(* IEC 61131-3 sources: Caravan/Archiv/12-04-19/Stations/MachineControl/MachineControl/Class/VaranManager (part 3) *)

#ifndef VARAN_TIME_MEASUREMENT_DEACTIVATE
        if pMultiVaran^.udVersion >= VM_MULTIVARAN_VERSION_FULL_PAYLOAD_AVAILABLE then
          //save max response time
          if ( p_node_info^^.uiResponseTimeMax > s_VaranTimes.ud_MaxResponseTime ) then

            s_VaranTimes.ud_MaxResponseTime := p_node_info^^.uiResponseTimeMax;

            //set T3 (no command executed before isochronous task)
            s_ManagerControlData.ud_MaxTimeCmdExecution := s_ManagerControlData.ud_IsoStartPoint -
                                  (2*( ( ( 276 * VM_TIMEOUT_ONE_BYTE )			//max 128 read/write befehl
                                    + s_VaranTimes.ud_MaxResponseTime       //The Manager need 2 Commands before he is free ( Prefetch + actual Command), reason for the whole term multiple 2
                                    )                                       //minimize the Jitter from the VARAN-BUS
                                    * ( VM_ALLOWED_RETRIES + 1 ))
                                  );

            //if time is neg set to 0
            if ( s_ManagerControlData.ud_MaxTimeCmdExecution$DINT < 0 ) then
              s_ManagerControlData.ud_MaxTimeCmdExecution := 0;
            end_if;

            // Write the data
            nodeProperty.udPropertyId    := VM_PROP_MAX_COMMAND_EXECUTION_TIME;
            nodeProperty.udPropertyValue := s_ManagerControlData.ud_MaxTimeCmdExecution;
            MULTI_VARAN_iSetNodeProperties( hNodeHandle           := vmNodeHandle
                                          , udPropertyCount       := 1
                                          , psPropertyValuePairs  := #nodeProperty
                                          );

          end_if;

        else
          //save max response time
          if ( p_node_info^^.uiResponseTimeMax > s_VaranTimes.ud_MaxResponseTime ) & p_ManagerStructure then

            s_VaranTimes.ud_MaxResponseTime := p_node_info^^.uiResponseTimeMax;

            //set T3 (no command executed before isochronous task)
            p_ManagerStructure^.uiMaxTimeCmdExecution := 	p_ManagerStructure^.uiIsoStartPoint -
                                  (2*( ( ( 276 * VM_TIMEOUT_ONE_BYTE )			//max 128 read/write befehl
                                    + s_VaranTimes.ud_MaxResponseTime       //The Manager need 2 Commands before he is free ( Prefetch + actual Command), reason for the whole term multiple 2
                                    )                                       //minimize the Jitter from the VARAN-BUS
                                    * ( VM_ALLOWED_RETRIES + 1 ))
                                  );

            //if time is neg set to 0
            if ( p_ManagerStructure^.uiMaxTimeCmdExecution$DINT < 0 ) then
              p_ManagerStructure^.uiMaxTimeCmdExecution := 0;
            end_if;
          end_if;
        end_if;
#endif

      else
        sd_retval := VM_CMD_ERROR_EMPTY_POINTER;
      end_if;

    elsif pVaran then  // if b_PayloadSupport then //----------------------------------------------------------------------------------------------------------

      //call OS - function to right device address
      sd_retval := VARAN_iGetNodeInfo	( uiManager	:= VaranManagerNr
                                      , pucNode	  := p_us_position_info
                                      , pNodeInfo	:= p_node_info
                                      );

      //look for an Error
      if ( sd_retval <> VARANMANAGER_OK ) then
        s_ErrorVaranManager.f_GetNodeInfo := SetVaranDOError( sd_Error 		  := sd_retval
                                                            , b_manager_off	:= FALSE
                                                            , b_log			    := FALSE
                                                            );
        return;
      end_if;

#ifndef VARAN_TIME_MEASUREMENT_DEACTIVATE
      //save max response time
      if ( p_node_info^^.uiResponseTimeMax > s_VaranTimes.ud_MaxResponseTime ) & p_ManagerStructure then

        s_VaranTimes.ud_MaxResponseTime := p_node_info^^.uiResponseTimeMax;

        //set T3 (no command executed before isochronous task)
        p_ManagerStructure^.uiMaxTimeCmdExecution := 	p_ManagerStructure^.uiIsoStartPoint -
                              (2*( ( ( 276 * VM_TIMEOUT_ONE_BYTE )			//max 128 read/write befehl
                                + s_VaranTimes.ud_MaxResponseTime       //The Manager need 2 Commands before he is free ( Prefetch + actual Command), reason for the whole term multiple 2
                                )                                       //minimize the Jitter from the VARAN-BUS
                                * ( VM_ALLOWED_RETRIES + 1 ))
                              );

        //if time is neg set to 0
        if ( p_ManagerStructure^.uiMaxTimeCmdExecution$DINT < 0 ) then
          p_ManagerStructure^.uiMaxTimeCmdExecution := 0;
        end_if;
      end_if;
#endif
    end_if;	  // if b_PayloadSupport then //----------------------------------------------------------------------------------------------------------

  else
    sd_retval := -101;
  end_if;

END_FUNCTION //VIRTUAL GLOBAL VaranManager::GetNodeInfo

//[#ENGLISH]
//=================================================================================================
//Function to get Varan Manager number
//=================================================================================================
//[clients]	VaranManagerNr		:R		:number of varan manager
//[members]	pVaran					:R		:pointer to varan os functions
//			s_VaranManagerSettings	:R		:structure for different varan settings
//[<sd_Manager_number]number of varan Manager
//[>p_varan]address of pointer to varan
FUNCTION VIRTUAL GLOBAL VaranManager::GetManagerNumber
  VAR_INPUT
    p_varan				    : ^pVoid;
  END_VAR
  VAR_OUTPUT
    ud_manager_number	:  UDINT;
  END_VAR

  //look if init was executed
  if ( s_VaranManagerSettings.us_InitCounter = 0 ) then
    bExternalInit := true;
    Init();
  end_if;

  //set pointer to varan functions
  p_varan^:= pVaran;

  //give back varan manager number
  ud_manager_number := VaranManagerNr.read();

END_FUNCTION //VIRTUAL GLOBAL VaranManager::GetManagerNumber

//[#ENGLISH]
//=================================================================================================
//Function to log faults in cyclic (to prevent an error 67)
//=================================================================================================
//[server]	State					:W		:State of class
//[members]	s_VaranManagerSettings	:W		:structure for different varan settings
FUNCTION  VaranManager::LogError
  VAR
    ud_reason	      : UDINT;
    b_SetError    	: BOOL;
  END_VAR

  ud_reason := 0;

  b_SetError := FALSE;

  //look which entry
  case ( State ) of
//**********************************************************************************************************************************************************
    _TimeSliceError:	//Log entry
#ifdef HWC_LogError
      HWC_LogError(this, "@06B8 (VaranManager::LogError) Timeslice Error! Manager is set off!");
#endif
      ud_reason := VM_ERROR_TIMESLICE;
      b_SetError := TRUE;

//**********************************************************************************************************************************************************
    _TimesliceErrorIRQ:	//Log entry
#ifdef HWC_LogError
      HWC_LogError(this, "@06C2 (VaranManager::LogError) Timeslice Error Interrupt, Manager is set off!");
#endif
      ud_reason := VM_ERROR_TIMESLICE_IRQ;
      b_SetError := TRUE;

//**********************************************************************************************************************************************************
    _WatchdogError:		//Log entry
#ifdef HWC_LogError
      HWC_LogError(this, "@06CC (VaranManager::LogError) Watchdog Error Interrupt, Manager is set off!");
#endif
      ud_reason := VM_ERROR_WATCHDOG;
      b_SetError := TRUE;

//**********************************************************************************************************************************************************
    _RequiredError:		//Log entry
#ifdef HWC_LogError
      HWC_LogError(this, "@06D6 (VaranManager::LogError) Required Module not ready, Manager is set off!");
#endif
      //b_SetError := FALSE;

//**********************************************************************************************************************************************************
    _DeviceError:		//Log entry
#ifdef HWC_LogError
      HWC_LogError(this, "@06E0 (VaranManager::LogError) Error on Device, Manager is set off!");
#endif
      ud_reason := VM_ERROR_DEVICE;
      b_SetError := TRUE;

//**********************************************************************************************************************************************************
    _CDIASRequiredError, _DIASRequiredError, _DiasError: //Log Entry
#ifdef HWC_LogError
      HWC_LogError(this, "@0024 (VaranManager::LogError) Required DIAS/CDIAS Module not ready, Manager is set off!");
#endif
      ud_reason   := VM_ERROR_DEVICE;
      b_SetError  := TRUE;
      State       := _RequiredError;

//**********************************************************************************************************************************************************
  else     //Unknown fault, log that an error occured
#ifdef HWC_LogValue1
    HWC_LogValue1(this, "@0025 (VaranManager::LogError) Unknown Fault (State = {0}), Manager is set off!", State);
#endif
  end_case;

  //reset log flag
  s_VaranManagerSettings.b_LogError := FALSE;

  //set Hw off
  To_HwControl.SetHardwareOff( e_error := State );

  //produce Varan Manager Error
  if ( b_SetError & PreventManagerError = 0) then

    if b_PayloadSupport & pMultiVaran^.udVersion >= VM_MULTIVARAN_VERSION_FULL_PAYLOAD_AVAILABLE  then
      MULTI_VARAN_iReportVaranError(diErrorNumber := ud_reason$DINT
                                  , hErrorNode    := vmNodeHandle);

    elsif pVaran & (pVaran^.udVersion >= 16#00001104 ) then
      VARAN_iSetManagerError( VaranManagerNr, ud_reason );
    end_if;
  end_if;

END_FUNCTION // VaranManager::LogError

//[#ENGLISH]
//=================================================================================================
//Function returns state of Varan manger class
//=================================================================================================
//[<e_state]error of varan manager
FUNCTION VIRTUAL GLOBAL VaranManager::GetManagerState
  VAR_OUTPUT
    e_state		  : t_e_VaranErrors;
  END_VAR

  e_state := State;

END_FUNCTION //VIRTUAL GLOBAL VaranManager::GetManagerState

//[#ENGLISH]
//=================================================================================================
//Function to add a multiple read/write register
//=================================================================================================
//[>p_us_position_info]pointer to position info( first byte is length)
//[>ud_dol_type] type of DOL list( 1=direct access, 2=IRQ, 3=realtime, 4=cyclic )
//[>p_ud_handle] pointer to variable to set right handle
//[>ud_address_read] Address of read data object
//[>ud_length_read] Length of read data object
//[>p_ud_data_read] pointer to variable to get pointer to data
//[>ud_address_write] Address of write data object
//[>ud_length_write] Length of write data object
//[>p_ud_data_write] pointer to variable to get pointer to data
//[>us_filter]filter number
//[>ui_number_of_slices]maximal number of slices
//[<sd_retval] 0=OK, negative=error (look lsl_st_varan.h)
FUNCTION GLOBAL VaranManager::AddMultipleRdWr
  VAR_INPUT
    p_us_position_info		: ^USINT;
    ud_dol_type				    :  UDINT;
    p_ud_handle				    : ^UDINT;
    ud_address_read			  :  UDINT;
    ud_length_read			  :  UDINT;
    p_ud_data_read			  : ^UDINT;
    ud_address_write		  :  UDINT;
    ud_length_write			  :  UDINT;
    p_ud_data_write			  : ^UDINT;
    us_filter				      :  USINT;
    ui_number_of_slices		:  UINT;
  END_VAR
  VAR_OUTPUT
    sd_retval				      :  DINT;
  END_VAR
  VAR
    ud_command			      :  UDINT;
    TempMem               :  UDINT;
  END_VAR

  //look if right OS - Version
  if ( _RTOSVersion >= 16#1194 ) & pVaran then

    //set command
    ud_command := VARAN_CMD_MULTIPLE_MEMORY_RW or ( us_filter shl 8 ) or ( ui_number_of_slices shl 16 );

    //look if we must execute Cyclic DOL list
    if ( ud_dol_type = VARAN_DOL_ASY ) then
      s_CyHandles.b_ExecuteDOL := TRUE;			//set flag to execut Dol list
    end_if;

    //Install Varan data object
    sd_retval := VARAN_iAddDOToDOL( uiManager     := VaranManagerNr
                                  , pucNode       := p_us_position_info
                                  , uiDOLType     := ud_dol_type
                                  , puiDOHandle   := p_ud_handle
                                  , uiCmd				  := ud_command
                                  , uiAddressRead := ud_address_read
                                  , uiLengthRead  := ud_length_read
                                  , pucRead       := p_ud_data_read
                                  , uiAddressWrite:= ud_address_write
                                  , uiLengthWrite := ud_length_write
                                  , pucWrite      := p_ud_data_write
                                  );

    //look if an error occured
    if ( sd_retval <> VARANMANAGER_OK ) then
      s_ErrorVaranManager.f_AddRdWrDO := SetVaranDOError( sd_Error      := sd_retval
                                                        , b_manager_off := TRUE
                                                        , b_log         := TRUE
                                                        );
    else
    //   32Byte (Header) +
    // + 13 Byte (Addr + Len +... --> See design spec appendix) +
    // + (1 Byte (Response) + n Byte) * slices (load data read) +
    // + n * slices Byte (load data write) +
    // + 0 to 3 Byte (compensate missalignment)
      TempMem := 32 + 13 + (1 + ud_length_read) * ui_number_of_slices + ud_length_write * ui_number_of_slices;
      if (TempMem MOD 4) then
        TempMem := TempMem + (4 - (TempMem MOD 4)); //increase memory, up to a value, which could be divided by 4
      end_if;

      if ud_dol_type = VARAN_DOL_ISO then
        DPRAM_Used.ISO_RdWr += TempMem;
        DOCounter.ISO_RdWr  += 1;
      else
        DPRAM_Used.ASY_RdWr += TempMem;
        DOCounter.ASY_RdWr  += 1;
      end_if;

      DPRAM_Used.Total      += TempMem;
      DOCounter.Total       += 1;
    end_if;
  else
    sd_retval := -100;	//Manager is off
  end_if;

END_FUNCTION //VIRTUAL GLOBAL VaranManager::AddMultipleRdWr

//[#ENGLISH]
//=================================================================================================
//Function to get an actual filter number
//=================================================================================================
//[<us_filter]number of filter
FUNCTION GLOBAL VaranManager::GetFilterNumber
  VAR_OUTPUT
    us_filter : USINT;
  END_VAR

  if ( s_VaranManagerSettings.us_FilterNumber <> 255 ) then
    //increment filter number
    s_VaranManagerSettings.us_FilterNumber += 1;
    us_filter := s_VaranManagerSettings.us_FilterNumber;
  else
    us_filter := 0;
  end_if;

END_FUNCTION //VIRTUAL GLOBAL VaranManager::GetFilterNumber

//[#ENGLISH]
//=================================================================================================
//Function to write a direct access data object
//=================================================================================================
//[members]	s_DirectAccessDO	:W/R	:structure for direct access
//[>p_us_position_info]pointer to position info( first byte is length)
//[>ud_address_read] Address of read data object
//[>ud_length_read] Length of read data object
//[>p_ud_data_read] pointer to variable to get pointer to data
//[>ud_address_write] Address of write data object
//[>ud_length_write] Length of write data object
//[>p_ud_data_write] pointer to variable to get pointer to data
//[>us_filter] number of filter
//[>us_slices] max number of slices
//[>p_handle]pointer to varan header
//[<sd_retval] 0=OK, negative=error (look lsl_st_varan.h)
FUNCTION GLOBAL VaranManager::MultipleRdWrDO
  VAR_INPUT
    p_us_position_info	: ^USINT;
    ud_address_read		  :  UDINT;
    ud_length_read		  :  UDINT;
    p_ud_data_read		  : ^UDINT;
    ud_address_write  	:  UDINT;
    ud_length_write		  :  UDINT;
    p_ud_data_write	  	: ^UDINT;
    us_filter			      :  USINT;
    us_slices			      :  USINT;
    p_handle			      : ^PLSL_VARANFRAME;
  END_VAR
  VAR_OUTPUT
    sd_retval		      	:  DINT;
  END_VAR

  //look if right OS - Version
  if ( _RTOSVersion >= 16#1194 ) then

    //clear direct access dol list
    sd_retval := ClearDOL( ud_dol_type := VARAN_DOL_DA );

    //look if an error occurs
    if ( sd_retval <> VARANMANAGER_OK ) then
      s_ErrorVaranManager.f_WrDO := SetVaranDOError	( sd_Error 	    := sd_retval
                                                    , b_manager_off	:= TRUE
                                                    , b_log			    := FALSE
                                                    );
      return;
    end_if;

    //add data object
    sd_retval := AddMultipleRdWr( p_us_position_info	:= p_us_position_info
                                , ud_dol_type			    := VARAN_DOL_DA
                                , p_ud_handle			    := p_handle$^UDINT
                                , ud_address_read		  := ud_address_read
                                , ud_length_read		  := ud_length_read
                                , p_ud_data_read		  := ( #p_ud_data_read )$^UDINT
                                , ud_address_write		:= ud_address_write
                                , ud_length_write		  := ud_length_write
                                , p_ud_data_write		  := ( #p_ud_data_write )$^UDINT
                                , us_filter				    := us_filter
                                , ui_number_of_slices	:= us_slices
                                );

    //look if an error occurs
    if ( sd_retval <> VARANMANAGER_OK ) then
      s_ErrorVaranManager.f_WrDO := SetVaranDOError	( sd_Error 		  := sd_retval
                                                    , b_manager_off	:= TRUE
                                                    , b_log			    := FALSE
                                                    );
      return;
    end_if;

    //set run status of data object on
    p_handle^^.ucCtrlStat 	        := VARAN_DO_SINGLE_RUN;

    //set number of allowed retries
    p_handle^^.ucRetrys	          	:= VM_ALLOWED_RETRIES;

    //set time for retry timeout
    p_handle^^.uiRetryTimeout       := VM_MAX_RETRY_TIMEOUT_MULTIPLE;

    //Execute dol
    sd_retval := ExecuteDOL( ud_dol_type := VARAN_DOL_DA );//or VARAN_DOL_EXECUTE_WAIT );

    //look if an error occurs
    if ( sd_retval <> VARANMANAGER_OK ) then
      s_ErrorVaranManager.f_WrDO := SetVaranDOError	( sd_Error 		  := sd_retval
                                                    , b_manager_off	:= TRUE
                                                    , b_log			    := FALSE
                                                    );
      return;
    end_if;

  else
    sd_retval := -100;	//Manager is off
  end_if;

END_FUNCTION //VIRTUAL GLOBAL VaranManager::MultipleRdWrDO

//[#ENGLISH]
//=================================================================================================
//Function to read SPI data
//=================================================================================================
//[>p_us_position_info]pointer to position info( first byte is length)
//[>ud_offset]offset in SPI flash
//[>ud_length]length of data (max. 128Byte)
//[>p_data]pointer to allocated memory for read data
//[<sd_retval] 0=OK, negative=error (look lsl_st_varan.h)
FUNCTION VIRTUAL GLOBAL VaranManager::ReadSPIData
  VAR_INPUT
    p_us_position_info	  : ^USINT;
    ud_offset		        	:  UDINT;
    ud_length		        	:  UDINT;
    p_data			        	: ^USINT;
  END_VAR
  VAR_OUTPUT
    sd_retval		          :  DINT;
  END_VAR
  VAR
    ud_sent_page	        :  UDINT;
    ud_NodeHandle         : UDINT;
    sPropertyValuePair    : LSL_PROPERTY_VALUE_PAIR;
  END_VAR

  //look if right OS - Version
  if ( _RTOSVersion >= 16#119F ) then

    if ( ud_length and VM_SPI_IDENT_LIST ) then
      ud_length     := ud_length and 16#7FFF_FFFF;
      ud_sent_page  := 16#FFFF_FFFF;   // = Read from the last page
    else
      ud_sent_page  := ud_offset / VM_SPI_PAGE_SIZE;
    end_if;

    //look for length
    if ( ud_length <= 0 | ud_length > 128 | p_data = NIL ) then
      sd_retval := -101;
      return;
    end_if;

    if b_PayloadSupport then
      // Get Node Handle
      sd_retval := MULTI_VARAN_iGetNodeHandle ( udManagerNumber := VaranManagerNr
                                              , pszHardwarePath := p_us_position_info
                                              , phNodeHandle    := #ud_NodeHandle
                                              );

      if sd_retval <> VARANMANAGER_OK then
        return;
      end_if;

      // set request
      sPropertyValuePair.udPropertyId     := ND_PROP_SPI_MASTER_REQUEST;
      sPropertyValuePair.udPropertyValue  := SPI_MASTER_REQ_SET;
      sd_retval := MULTI_VARAN_iSetNodeProperties ( hNodeHandle           := ud_NodeHandle
                                                  , udPropertyCount       := 1
                                                  , psPropertyValuePairs  := #sPropertyValuePair
                                                  );
      // look for an error
      if ( sd_retval <> VARANMANAGER_OK ) then
        return;
      end_if;

      // set right page
      sd_retval := MULTI_VARAN_iSpiMasterReadFlashPage( hNodeHandle           := ud_NodeHandle
                                                      , udPageNumber          := ud_sent_page
                                                      , udOffsetInPage        := ud_offset mod VM_SPI_PAGE_SIZE
                                                      , udReadLength          := ud_length
                                                      , bBlockUntilCompleted  := true
                                                      , pusData               := p_data
                                                      );
      //look for an error
      if ( sd_retval <> VARANMANAGER_OK ) then
        return;
      end_if;

      //clear request
      sPropertyValuePair.udPropertyId     := ND_PROP_SPI_MASTER_REQUEST;
      sPropertyValuePair.udPropertyValue  := SPI_MASTER_REQ_CLEARED;
      sd_retval := MULTI_VARAN_iSetNodeProperties ( hNodeHandle           := ud_NodeHandle
                                                  , udPropertyCount       := 1
                                                  , psPropertyValuePairs  := #sPropertyValuePair
                                                  );
    elsif pVaran then

      //set request
    sd_retval := VARAN_iSPIMasterSetRequest	( uiManager	:= VaranManagerNr
                                            , pucNode	  := p_us_position_info
                                            );

    //look for an error
    if ( sd_retval <> VARANMANAGER_OK ) then
      return;
    end_if;

    //set right page
    sd_retval := VARAN_iSPIMasterPageRead	( uiManager	:= VaranManagerNr
                                          , pucNode	  := p_us_position_info
                                          , uiPage	  := ud_sent_page
                                          );

    //look for an error
    if ( sd_retval <> VARANMANAGER_OK ) then
      return;
    end_if;

    ud_sent_page := ud_offset mod VM_SPI_PAGE_SIZE;

    //read data of page
    sd_retval := VARAN_iSPIMasterPageReadBuffer	( uiManager	:= VaranManagerNr
                                                , pucNode	  := p_us_position_info
                                                , uiOffset	:= ud_sent_page
                                                , uiLen		  := ud_length
                                                , puiPage	  := p_data
                                                );

    //look for an error
    if ( sd_retval <> VARANMANAGER_OK ) then
      return;
    end_if;

    //clear request
    sd_retval := VARAN_iSPIMasterClearRequest	( uiManager	:= VaranManagerNr
                                              , pucNode	  := p_us_position_info
                                              );
    end_if;

  else
    sd_retval := -100;
  end_if;

END_FUNCTION //VIRTUAL GLOBAL VaranManager::ReadSPIData

//[#ENGLISH]
//=================================================================================================
//Function add a foreign package request
//=================================================================================================
//[>p_us_position_info]pointer to position info( first byte is length)
//[>ud_dol_type] type of DOL list( 1=direct access, 2=IRQ, 3=realtime, 4=cyclic )
//[>p_ud_handle]pointer to variable to set right handle
//[>ud_address] Address of data object
//[<sd_retval] 0=OK, negative=error (look lsl_st_varan.h)
FUNCTION VIRTUAL GLOBAL VaranManager::AddForeignPackRequest
  VAR_INPUT
    p_us_position_info	: ^USINT;
    ud_dol_type		    	: UDINT;
    p_ud_handle			    : ^UDINT;
    ud_address			    : UDINT;
  END_VAR
  VAR_OUTPUT
    sd_retval		      	: DINT;
  END_VAR
  VAR
    ud_NodeHandle       : UDINT;
  END_VAR

  //look if we must execute Cyclic DOL list
  if ( ud_dol_type = VARAN_DOL_ASY ) then
    s_CyHandles.b_ExecuteDOL := TRUE;			//set flag to execut Dol list
  end_if;

  if b_PayloadSupport &
       pMultiVaran^.udVersion >= VM_MULTIVARAN_VERSION_FULL_PAYLOAD_AVAILABLE  then
    sd_retval := MULTI_VARAN_iGetNodeHandle ( udManagerNumber := VaranManagerNr
                                            , pszHardwarePath := p_DisablePath
                                            , phNodeHandle    := #ud_NodeHandle
                                            );

    // Return the ErrorCode
    if sd_retval then
      return;
    end_if;

    sd_retval := MULTI_VARAN_iAddDo(  phDoHandle                    := p_ud_handle
                                    , hNodeHandle                   := ud_NodeHandle
                                    , bDoRequired                   := 0
                                    , udDolType                     := ud_dol_type
                                    , udCommand                     := VARAN_CMD_FOREIGN_PACKET_REQ
                                    , udPriority                    := VM_PRIORITY_READ_DO
                                    , udPrescalerCounterThreshold   := 0
                                    , udPrescalerCounterStartValue  := 0
                                    , udReadOffset                  := VARAN_CLIENT_FP_SAFETY
                                    , udReadLength                  := VARAN_FPR_SAFETY_ID
                                    , udWriteOffset                 := 0
                                    , udWriteLength                 := 0
                                    , udFilter                      := 0
                                    , udSlices                      := 0
                                    , udWritePayloadType            := WR_PLD_TYPE_STANDARD
                                    );

  else
    // if there is no VARAN Interface available, we would crash at the call
    if pVaran = NIL then
      sd_retval := VARANMANAGER_DRIVER_NOT_EXISTS;
      return;
    end_if;

    //Install Varan data object
    sd_retval := VARAN_iAddDOToDOL	( uiManager			  := VaranManagerNr
                                    , pucNode			    := p_us_position_info
                                    , uiDOLType 		  := ud_dol_type + ( VARAN_DO_EXECUTE_FIFO_EMPTY shl 24 ) // in the highest byte we have the init value for the uc_CtrlStat Register
                                    , puiDOHandle		  := p_ud_handle
                                    , uiCmd				    := VARAN_CMD_FOREIGN_PACKET_REQ
                                    , uiAddressRead		:= ud_address + VARAN_CLIENT_FP_SAFETY
                                    , uiLengthRead		:= VARAN_FPR_SAFETY_ID
                                    , pucRead			    := NIL
                                    , uiAddressWrite	:= 0
                                    , uiLengthWrite		:= 0
                                    , pucWrite			  := NIL
                                    );
  end_if;

  //look if an error occured
  if ( sd_retval <> VARANMANAGER_OK ) then
    s_ErrorVaranManager.f_AddFoPaReq := SetVaranDOError ( sd_Error 		  := sd_retval
                                                        , b_manager_off	:= TRUE
                                                        , b_log			    := TRUE
                                                        );
  end_if;

  //look if an error occured
  if ( sd_retval <> VARANMANAGER_OK ) then
    s_ErrorVaranManager.f_AddFoPaReq := SetVaranDOError ( sd_Error 		  := sd_retval
                                                        , b_manager_off	:= TRUE
                                                        , b_log			    := TRUE
                                                        );
  end_if;

END_FUNCTION //VIRTUAL GLOBAL VaranManager::AddForeignPackRequest

//[#ENGLISH]
//=================================================================================================
//Function to get sync frame counter
//=================================================================================================
//[<us_frame_counter] sync frame counter
FUNCTION VIRTUAL GLOBAL VaranManager::GetSyncFrameCounter
  VAR_OUTPUT
    us_frame_counter		: USINT;
  END_VAR

  if b_PayloadSupport &
     pMultiVaran^.udVersion >= VM_MULTIVARAN_VERSION_FULL_PAYLOAD_AVAILABLE  then
    MULTI_VARAN_iGetNodeProperty( hNodeHandle       := vmNodeHandle
                                , udPropertyId      := VM_PROP_SYNC_COUNTER
                                , pudPropertyValue  := (#us_frame_counter)$^UDINT
                                );
  else
    us_frame_counter := p_SyncData^.us_FrameCounter;
  end_if;

END_FUNCTION //VIRTUAL GLOBAL VaranManager::GetSyncFrameCounter

//[<retval]ISO start point [ns]
FUNCTION VIRTUAL GLOBAL VaranManager::GetIsoStartPoint
  VAR_OUTPUT
    retval	  	: UDINT;
  END_VAR

  //if init is not executed yet
  if ( s_VaranManagerSettings.us_InitCounter = 0 ) then
    GetISOStartTime();
  end_if;

  retval := VaranManagerTime * IsoStartPoint / 100;

END_FUNCTION //VIRTUAL GLOBAL VaranManager::GetIsoStartPoint

FUNCTION  VaranManager::GetISOStartTime

  //set realtime start point of varan list
  //VaranManagerTime must be below 47ms!
  IsoStartPoint := IsoStartPoint.Read();
  if( IsoStartPoint < 1 )then
    IsoStartPoint := 50;
  end_if;
  if( IsoStartPoint > 99 )then
    IsoStartPoint := 50;
  end_if;

END_FUNCTION // VaranManager::GetISOStartTime

//=================================================================================================
//Function to set disable device in cyclic
//=================================================================================================
//[>p_us_position_info]path of varan
FUNCTION VIRTUAL GLOBAL VaranManager::SetDisableDevice
  VAR_INPUT
    p_us_position_info		: ^USINT;
  END_VAR
  VAR_OUTPUT
    sd_retval		          :  DINT;
  END_VAR

  sd_retval := -100;

  if ( b_DisableDevice = FALSE ) then
    b_DisableDevice := TRUE;
    p_DisablePath   := p_us_position_info;
    sd_retval       := 0;
  end_if;

END_FUNCTION //VIRTUAL GLOBAL VaranManager::SetDisableDevice

//=================================================================================================
//Function to disable device in cyclic
//=================================================================================================
FUNCTION  VaranManager::DisableDevice
  VAR_OUTPUT
    sd_retval		    : DINT;
  END_VAR
  VAR
    ud_NodeHandle   : UDINT;
    nodeProperty    : LSL_PROPERTY_VALUE_PAIR;
  END_VAR

  if b_PayloadSupport &
     pMultiVaran^.udVersion > VM_MULTIVARAN_VERSION_FULL_PAYLOAD_AVAILABLE then

    sd_retval := MULTI_VARAN_iGetNodeHandle ( udManagerNumber := VaranManagerNr
                                            , pszHardwarePath := p_DisablePath
                                            , phNodeHandle    := #ud_NodeHandle
                                            );

    // Return the ErrorCode
    if sd_retval then
      return;
    end_if;

    nodeProperty.udPropertyId    := ND_PROP_CONNECTION_STATE;
    nodeProperty.udPropertyValue := CN_STATE_DISCONNECTED;
    sd_retval := MULTI_VARAN_iSetNodeProperties ( hNodeHandle           := ud_NodeHandle
                                                , udPropertyCount       := 1
                                                , psPropertyValuePairs  := #nodeProperty
                                                );

  //look if funtion is available with this os version
  elsif ( _RTOSVersion >= VM_DISABLE_DEVICE_AVAILABLE ) & pVaran then

    //disable device
    sd_retval := VARAN_iSetNodeEnableStatus	( uiManager		  := VaranManagerNr
                                            , pucNode		    := p_DisablePath
                                            , uiNodeStatus	:= 0
                                            );

    b_DisableDevice := FALSE;

  else
    sd_retval := -100;
  end_if;

END_FUNCTION // VaranManager::DisableDevice

FUNCTION GLOBAL VaranManager::ReadWaitingTimeBeforeSync
  VAR_OUTPUT
    ud_waitingtime 	  : UDINT;
  END_VAR

  ud_waitingtime := 0;

  if b_PayloadSupport  &
    pMultiVaran^.udVersion >= VM_MULTIVARAN_VERSION_FULL_PAYLOAD_AVAILABLE then

    ud_waitingtime := s_ManagerControlData.ud_IsoStartPoint - s_ManagerControlData.ud_MaxTimeCmdExecution;

  // check manager structure
  elsif ( p_ManagerStructure ) then
     ud_waitingtime := p_ManagerStructure^.uiIsoStartPoint - p_ManagerStructure^.uiMaxTimeCmdExecution;
  end_if;

END_FUNCTION

FUNCTION GLOBAL VaranManager::SetWaitingTimeBeforeSync
  VAR_INPUT
    ud_waitingtime 	: UDINT;
  END_VAR
  VAR
    nodeProperty    : LSL_PROPERTY_VALUE_PAIR;
  END_VAR

  if b_PayloadSupport  &
     pMultiVaran^.udVersion >= VM_MULTIVARAN_VERSION_FULL_PAYLOAD_AVAILABLE then
    //set T3 (no command executed before isochronous task)
    s_ManagerControlData.ud_MaxTimeCmdExecution := s_ManagerControlData.ud_IsoStartPoint - ud_waitingtime;

    //if time is neg set to 0
    if ( s_ManagerControlData.ud_MaxTimeCmdExecution$DINT < 0 ) then
      s_ManagerControlData.ud_MaxTimeCmdExecution := 0;
    end_if;

    // Write the data
    nodeProperty.udPropertyId    := VM_PROP_MAX_COMMAND_EXECUTION_TIME;
    nodeProperty.udPropertyValue := s_ManagerControlData.ud_MaxTimeCmdExecution;
    MULTI_VARAN_iSetNodeProperties( hNodeHandle           := vmNodeHandle
                                  , udPropertyCount       := 1
                                  , psPropertyValuePairs  := #nodeProperty
                                  );

  elsif ( p_ManagerStructure ) then

    //set T3 (no command executed before isochronous task)
    p_ManagerStructure^.uiMaxTimeCmdExecution := 	p_ManagerStructure^.uiIsoStartPoint - ud_waitingtime;

    //if time is neg set to 0
    if ( p_ManagerStructure^.uiMaxTimeCmdExecution$DINT < 0 ) then
      p_ManagerStructure^.uiMaxTimeCmdExecution := 0;
    end_if;
  end_if;

END_FUNCTION

FUNCTION VIRTUAL GLOBAL VaranManager::AddIsoClientRdData
  VAR_INPUT
    ud_length 	: UDINT;
    p_pdata 	  : ^void;
  END_VAR
  VAR_OUTPUT
    sd_retval 	: DINT;
  END_VAR

  if (IsAlsoClient <> 0) & (SuperiorSystemTime <> 0) then
    if us_InitCounter < 6 then
      if (SafetyIsoMemRead$UDINT + ud_length) <= (VM_CLIENT_MAX_BUFFER_USE - VM_CLIENT_HEADER_SIZE) then
        if p_pdata <> NIL then
          if UserObjectData.pIsoReadData = NIL then
            UserObjectData.udIsoReadLength := ud_length;
            UserObjectData.pIsoReadData    := p_pdata;
            sd_retval := 0;       // OK
          else
            sd_retval := -4;      // adding was allready done
          end_if;
        else
          sd_retval := -3;        // invalid pointer
        end_if;
      else
        sd_retval := -2;          // invalid length
      end_if;
    else
      sd_retval := -1;            // method was called to late
    end_if;
  else
    sd_retval := -5;              // wrong client settings
  end_if;

END_FUNCTION //GLOBAL VaranManager::AddIsoClientRdData

FUNCTION VIRTUAL GLOBAL VaranManager::AddIsoClientWrData
  VAR_INPUT
    ud_length 	: UDINT;
    p_pdata 	  : ^void;
  END_VAR
  VAR_OUTPUT
    sd_retval 	: DINT;
  END_VAR

  if (IsAlsoClient <> 0) & (SuperiorSystemTime <> 0) then
    if us_InitCounter < 6 then
      if (SafetyIsoMemWrite$UDINT + ud_length) <= (VM_CLIENT_MAX_BUFFER_USE - VM_CLIENT_HEADER_SIZE) then
        if p_pdata <> NIL then
          if UserObjectData.pIsoWriteData = NIL then
            UserObjectData.udIsoWriteLength := ud_length;
            UserObjectData.pIsoWriteData    := p_pdata;
            sd_retval := 0;       // OK
          else
            sd_retval := -4;      // adding was allready done
          end_if;
        else
          sd_retval := -3;        // invalid pointer
        end_if;
      else
        sd_retval := -2;          // invalid length
      end_if;
    else
      sd_retval := -1;            // method was called to late
    end_if;
  else
    sd_retval := -5;              // wrong client settings
  end_if;

END_FUNCTION //GLOBAL VaranManager::AddIsoClientWrData

FUNCTION VIRTUAL GLOBAL VaranManager::AddAsyClientRdData
  VAR_INPUT
    ud_length 	: UDINT;
    p_pdata 	  : ^void;
  END_VAR
  VAR_OUTPUT
    sd_retval 	: DINT;
  END_VAR

  if (IsAlsoClient <> 0) & (SuperiorSystemTime <> 0) then
    if us_InitCounter < 6 then
      if (SafetyAsyMemRead$UDINT + ud_length) <= (VM_CLIENT_MAX_BUFFER_USE - VM_CLIENT_HEADER_SIZE) then
        if p_pdata <> NIL then
          if UserObjectData.pAsyReadData = NIL then
            UserObjectData.udAsyReadLength  := ud_length;
            UserObjectData.pAsyReadData     := p_pdata;
            sd_retval := 0;       // OK
          else
            sd_retval := -4;      // adding was allready done
          end_if;
        else
          sd_retval := -3;        // invalid pointer
        end_if;
      else
        sd_retval := -2;          // invalid length
      end_if;
    else
      sd_retval := -1;            // method was called to late
    end_if;
  else
    sd_retval := -5;              // wrong client settings
  end_if;

END_FUNCTION //GLOBAL VaranManager::AddASYClientRdData

FUNCTION VIRTUAL GLOBAL VaranManager::AddAsyClientWrData
  VAR_INPUT
    ud_length 	: UDINT;
    p_pdata 	  : ^void;
  END_VAR
  VAR_OUTPUT
    sd_retval 	: DINT;
  END_VAR

  if (IsAlsoClient <> 0) & (SuperiorSystemTime <> 0) then
    if us_InitCounter < 6 then
      if (SafetyAsyMemWrite$UDINT + ud_length) <= (VM_CLIENT_MAX_BUFFER_USE - VM_CLIENT_HEADER_SIZE) then
        if p_pdata <> NIL  then
          if UserObjectData.pAsyWriteData = NIL then
            UserObjectData.udAsyWriteLength := ud_length;
            UserObjectData.pAsyWriteData    := p_pdata;
            sd_retval := 0;       // OK
          else
            sd_retval := -4;      // adding was allready done
          end_if;
        else
          sd_retval := -3;        // invalid pointer
        end_if;
      else
        sd_retval := -2;          // invalid length
      end_if;
    else
      sd_retval := -1;            // method was called to late
    end_if;
  else
    sd_retval := -5;              // wrong client settings
  end_if;

END_FUNCTION //GLOBAL VaranManager::AddASYClientWrData

FUNCTION VaranManager::ActISOReadLength
  VAR_INPUT
    loop 	  : USINT;
  END_VAR
  VAR_OUTPUT
    length 	: UDINT;
  END_VAR

  if (loop + 1) < ISORdVaranPackages then
    length := 128;
    return;
  end_if;

  if (loop + 1) = ISORdVaranPackages then
    length := ISOLastPackageRdSize;
  else
    length := 0;
  end_if;

END_FUNCTION

FUNCTION VaranManager::ActISOWriteLength
  VAR_INPUT
    loop 	  : USINT;
  END_VAR
  VAR_OUTPUT
    length 	: UDINT;
  END_VAR

  if (loop + 1) < ISOWrVaranPackages then
    length := 128;
    return;
  end_if;

  if (loop + 1) = ISOWrVaranPackages then
    length := ISOLastPackageWrSize;
  else
    length := 0;
  end_if;

END_FUNCTION

FUNCTION VaranManager::ActASYReadLength
  VAR_INPUT
    loop 	  : USINT;
  END_VAR
  VAR_OUTPUT
    length 	: UDINT;
  END_VAR

  if (loop + 1) < ASYRdVaranPackages then
    length := 128;
    return;
  end_if;

  if (loop + 1) = ASYRdVaranPackages then
    length := ASYLastPackageRdSize;
  else
    length := 0;
  end_if;

END_FUNCTION

FUNCTION VaranManager::ActASYWriteLength
  VAR_INPUT
    loop 	  : USINT;
  END_VAR
  VAR_OUTPUT
    length 	: UDINT;
  END_VAR

  if (loop + 1) < ASYWrVaranPackages then
    length := 128;
    return;
  end_if;

  if (loop + 1) = ASYWrVaranPackages then
    length := ASYLastPackageWrSize;
  else
    length := 0;
  end_if;

END_FUNCTION

FUNCTION VaranManager::InitMulDivVMC
  VAR_OUTPUT
    sd_retval 	: DINT;
  END_VAR
  VAR
    i           : DINT;
    Divi        : USINT;
    VaranMulti  : USINT;
    CPUMulti    : USINT;
    nodeProperty: ARRAY [0..2] OF LSL_PROPERTY_VALUE_PAIR;
  END_VAR

  // initialize return value
  sd_retval := 0;

  //set right pointer
  p_ManagerClientSpace$UDINT += VM_CLIENT_OFFSET;

  //superior time must not zero
  if ( SuperiorSystemTime = 0 ) then
    State := _VaranTimeError;
    IF ( _firstscan = TRUE ) THEN
      //Log entry
#ifdef HWC_LogError
      HWC_LogError(this, "@06EA (VaranManager::InitMulDivVMC) SuperiorSystemTime is 0!");
#endif
    END_IF;
    sd_retval := -1;
    return;
  end_if;

  if b_PayloadSupport &
     pMultiVaran^.udVersion >= VM_MULTIVARAN_VERSION_FULL_PAYLOAD_AVAILABLE  then  // -------------------------------------------------------------------

    // Sync outs are no longer written with DA, changes are stored locally and writte once
    p_SyncOutISOSwitch := #s_SyncOutISOSwitch;

  else  // if b_PayloadSupport then  // -------------------------------------------------------------------

    //look for right sync out pointer
    p_SyncOutISOSwitch := #p_ManagerPll^.sSynOutPeripheral1;

    //look in all peripheral sync outs
    for i := 1 to VM_MAX_SYNC_OUTS - 1 do

      //look if sync out id is correct
      if ( p_SyncOutISOSwitch^.ucSyncOutID = VM_CLIENT_ISO_SWITCH_ID ) then
        exit;					//we found right sync out --> exit
      end_if;

      //get pointer to next sync out
      p_SyncOutISOSwitch += sizeof ( LSL_VARANPLLSYNCOUT );

      //if we searched all sync outs without success, leave method
      if ( i = VM_MAX_SYNC_OUTS - 1 ) then
        //Log entry
#ifdef HWC_LogError
        HWC_LogError(this, "@06F4 (VaranManager::InitMulDivVMC) Couldn't find sync out for switching alternating buffer");
#endif

        State     := _PllError;
        sd_retval := -2;
        return;
      end_if;
    end_for;
  end_if; // if b_PayloadSupport then  // -------------------------------------------------------------------

  // check if the varan times are multiple of each other
  if ((VaranManagerTime MOD SuperiorSystemTime) <> 0) &
     ((SuperiorSystemTime MOD VaranManagerTime) <> 0) then

    //Log entry
#ifdef HWC_LogError
    HWC_LogError(this, "@06FE (VaranManager::InitMulDivVMC) VaranTime of superior system and inferior system have to be multiples of each other");
#endif

    State     := _PllError;
    sd_retval := -3;
    return;
  end_if;

  // check if the superior varan time is multiple of inferior system time
  if ((MainTimer MOD SuperiorSystemTime) <> 0) &
     ((SuperiorSystemTime MOD MainTimer) <> 0) then

    //Log entry
#ifdef HWC_LogError
    HWC_LogError(this, "@0708 (VaranManager::InitMulDivVMC) VaranTime of superior system and maintimer of inferior system have to be multiples of each other");
#endif

    State     := _PllError;
    sd_retval := -4;
    return;
  end_if;

  // check factor of superior varan time to inferior system time (maintimer)
  if (MainTimer <= SuperiorSystemTime) then
    // if system cycle times are different (master is slower), calculate difference (rounded)
    CPUMulti  := 1;
    Divi      := to_usint(SuperiorSystemTime / MainTimer);
    if (Divi < 1) then
      Divi := 1;
    end_if;
  else
    // if system cycle times are different (slave is slower), calculate difference (rounded)
    Divi := 1;
    CPUMulti := to_usint(MainTimer / SuperiorSystemTime);
    if (CPUMulti < 1) then
      CPUMulti := 1;
    end_if;
  end_if;

  if b_PayloadSupport &
     pMultiVaran^.udVersion >= VM_MULTIVARAN_VERSION_GET_SYSTEM_PROPERTY_AVAILABLE  then
    // Bit settig is done be the OS
    // set System Period Time
    nodeProperty[0].udPropertyId    := VM_PROP_PLL_SYSTEM_PERIOD_TIME;
    nodeProperty[0].udPropertyValue := SuperiorSystemTime / 10;

    // set System Period Divider (Pll)
    nodeProperty[1].udPropertyId    := VM_PROP_PLL_SYSTEM_PERIOD_DIVIDER;
    nodeProperty[1].udPropertyValue := Divi;

    MULTI_VARAN_iSetNodeProperties( hNodeHandle           := vmNodeHandle
                                  , udPropertyCount       := 2
                                  , psPropertyValuePairs  := #nodeProperty[0]);

    // if slave is slower and OS would be slower than 1ms because sync input, we use multiplier for CPU also
    if (SuperiorSystemTime < 1000000) & (CPUMulti > 1) then
      MULTI_VARAN_ICONFIGUREPLLSYNCOUT( hManagerNodeHandle    := vmNodeHandle
                                      , udSyncOutId           := VM_SYNC_CPU_ID
                                      , udPeriodMultiplier    := CPUMulti
                                      , udFrameCountThreshold := 0
                                      , udControlStatus       := 1
                                      );  // enable cpu sync out in any case and enable frame count
    else
      MULTI_VARAN_ICONFIGUREPLLSYNCOUT( hManagerNodeHandle    := vmNodeHandle
                                      , udSyncOutId           := VM_SYNC_CPU_ID
                                      , udPeriodMultiplier    := 1
                                      , udFrameCountThreshold := 0
                                      , udControlStatus       := 1
                                      );  // enable cpu sync out in any case and enable frame count
    end_if;

  else

  // disable divider (bit 4) and pll (bit 6)
  p_ManagerPll^.ucControlStatus := p_ManagerPll^.ucControlStatus and 2#10101111;

  // set System Period Time
  p_ManagerPll^.aucPeriod$UDINT := SuperiorSystemTime / 10;

  // set System Period Divider (Pll)
  p_ManagerPll^.ucSystemPeriodDivider := Divi; // if you get an error on this line, you need the new lsl_st_varan.h where the name of the structure element is corrected

  // enable divider (bit 4) and pll (bit 6)
  p_ManagerPll^.ucControlStatus := p_ManagerPll^.ucControlStatus or 2#01010000;

  // if slave is slower and OS would be slower than 1ms because sync input, we use multiplier for CPU also
  if (SuperiorSystemTime < 1000000) & (CPUMulti > 1) then
    p_ManagerPll^.sSynOutCPU.ucPeriodMultiplier   := CPUMulti;
  else
    p_ManagerPll^.sSynOutCPU.ucPeriodMultiplier   := 1;
  end_if;
  p_ManagerPll^.sSynOutCPU.ucFrameCountThreshold  := 0;
  p_ManagerPll^.sSynOutCPU.ucControlStatus        := 1; // enable cpu sync out in any case and enable frame count
  end_if;

  VaranMulti := to_usint(VaranManagerTime / MainTimer) * CPUMulti;

  // get modulo value for synchronity check
  if SuperiorSystemTime > VaranManagerTime then
    VMC_ModValue := SuperiorSystemTime / VaranManagerTime;
    if VMC_ModValue < 1 then
      VMC_ModValue := 1;
    end_if;
  else
    VMC_ModValue := 1;
  end_if;

  // set Period Multiplier of Varan Manager
  p_SyncOut^.ucPeriodMultiplier := VaranMulti;

  ucVaranManagerTemp := 2#011; // framecounter

  // enable iso switch sync (bit0 = 1) in RtWork together with varan sync
  if (VaranMulti > 1) then
    // set Period Multiplier of ISO Switch
    p_SyncOutISOSwitch^.ucPeriodMultiplier := VaranMulti;

    // if (divisor > 1) and (superior time is not greater) then use system sync of superior system
    if (Divi > 1) & (SuperiorSystemTime <= VaranManagerTime) then
      ucVaranManagerTemp  :=
      ucIsoSwitchTemp     := 2#101;

      // correct multipliers
      p_SyncOutISOSwitch^.ucPeriodMultiplier  /= Divi;
      p_SyncOut^.ucPeriodMultiplier           /= Divi;
    else
      // if superior time is greater use superior sync for iso switch
      if (SuperiorSystemTime > VaranManagerTime) then
        p_SyncOutISOSwitch^.ucPeriodMultiplier := 1;
        ucIsoSwitchTemp := 2#101;
      else
        // otherwise divided sync
        ucIsoSwitchTemp := 2#011; // framecounter
      end_if;
    end_if;
  else
    // set Period Multiplier of ISO Switch
    p_SyncOutISOSwitch^.ucPeriodMultiplier := 1;

    // use system sync of superior system (bit2 = 1)
    ucIsoSwitchTemp := 2#101;
  end_if;

  // Write p_SyncOutISOSwitch, (p_SyncOut is written at the end of FirstInit)
  if b_PayloadSupport  &
     pMultiVaran^.udVersion >= VM_MULTIVARAN_VERSION_FULL_PAYLOAD_AVAILABLE then
    MULTI_VARAN_ICONFIGUREPLLSYNCOUT( hManagerNodeHandle    := vmNodeHandle
                                    , udSyncOutId           := VM_CLIENT_ISO_SWITCH_ID
                                    , udPeriodMultiplier    := p_SyncOutISOSwitch^.ucPeriodMultiplier
                                    , udFrameCountThreshold := p_SyncOutISOSwitch^.ucFrameCountThreshold
                                    , udControlStatus       := p_SyncOutISOSwitch^.ucControlStatus
                                    );
  end_if;

END_FUNCTION

FUNCTION GLOBAL VaranManager::FrameCounterChanged
  VAR_INPUT
    pOld 	  : ^USINT;
    pAct 	  : ^USINT;
  END_VAR
  VAR_OUTPUT
    retcode : BOOL;
  END_VAR
  VAR
    Temp    : USINT;
  END_VAR

  if b_PayloadSupport &
     pMultiVaran^.udVersion >= VM_MULTIVARAN_VERSION_FULL_PAYLOAD_AVAILABLE  then
    MULTI_VARAN_iGetNodeProperty( hNodeHandle       := vmNodeHandle
                                , udPropertyId      := VM_PROP_PLL_SYNC_TIME_FRAME_COUNTER
                                , pudPropertyValue  := (#Temp)$^UDINT
                                );
  else
    Temp := p_ManagerPll^.ucSyncTimeFrameCounter;
  end_if;

  if pOld & pAct then
    pOld^ := OldFrameCounter;
    pAct^ := Temp;
  end_if;

  if Temp <> OldFrameCounter then
    retcode         := TRUE;
    OldFrameCounter := Temp;
  else
    retcode := FALSE;
  end_if;

END_FUNCTION

FUNCTION VIRTUAL GLOBAL VaranManager::GetDocumentation
  VAR_INPUT
    p_us_position_info 	: ^USINT;
    p_dpne 	            : ^CHAR;
  END_VAR
  VAR_OUTPUT
    sd_retval 	        : DINT;
  END_VAR
  VAR
    FileHandle          : DINT;
    FileData            : ^USINT;
    BaseListAddress     : UDINT;
  END_VAR

  sd_retval := 0;

  if p_us_position_info & p_dpne then

    // try to open file
    FileHandle := To_FileSys.FileOpen( filename   := p_dpne,
                                       attributes := ATT_CREATE_ALWAYS
                                     );

    // check success of opening file
    if FileHandle >= 0 then

      //check OS version
      if ( _RTOSVersion < VM_SPI_OS_VERSION ) then
        // access of SPI flash not possible
        sd_retval := -3;
        return;
      end_if;

      // check if documentation is available and get file size and offset in SPI flash
      if ( SearchSPIList(p_us_position_info, VM_SPI_DOCU_ID, #BaseListAddress) <> VARANMANAGER_OK ) then
        sd_retval := -4;
        return;
      end_if;

      sd_retval := GetDocuFileInfo(p_us_position_info := p_us_position_info,
                                   ud_listOffset      := BaseListAddress
                                  );

      //allocate memory for the file data
      FileData := ( To_StdLib.Malloc( size := ud_SPI_Docu_Length ) )$^USINT;

      if ( FileData = NIL ) then
        State := _MemoryFault;
        sd_retval := -5;
        return;
      end_if;

      //read the whole file
      sd_retval := ReadSPIDataComfort( p_us_position_info := p_us_position_info,
                                       ud_offset	        := ud_SPI_Offset,
                                       ud_length	        := ud_SPI_Docu_Length,
                                       p_data		          := FileData
                                     );
      //look for an error
      if ( sd_retval <> VARANMANAGER_OK ) then
        sd_retval := -6;
        return;
      end_if;

      // write bytes into file
      if To_FileSys.FileWrite( handle := FileHandle,
                               buffer := FileData,
                               length := ud_SPI_Docu_Length
                             ) <> ud_SPI_Docu_Length$DINT then
        sd_retval := -7;
      end_if;

      To_StdLib.Free(FileData);
      To_FileSys.FileClose(handle := FileHandle);
    else
      // failed to open file
      sd_retval := -2;
    end_if;
  else
    // invalid parameters
    sd_retval := -1;
  end_if;

END_FUNCTION

FUNCTION VaranManager::SearchSPIList
  VAR_INPUT
    p_us_position_info 	: ^USINT;
    SearchID 	          : UDINT;
    p_BaseListAddress   : ^UDINT;
  END_VAR
  VAR_OUTPUT
    sd_retval 	        : DINT;
  END_VAR
  VAR
    i				            : UDINT;
    a_data              : ARRAY[0..31] OF UDINT;
  END_VAR

  if p_BaseListAddress = NIL then
    // invalid parameters
    sd_retval := -101;
    return;
  end_if;

  //read SPI data
  sd_retval := ReadSPIData( p_us_position_info	:= p_us_position_info
                          , ud_offset				    := 0
                          , ud_length				    := 128 or VM_SPI_IDENT_LIST
                          , p_data				      := ( #a_data )$^USINT
                          );

  //look for an error
  if ( sd_retval <> VARANMANAGER_OK ) then
    return;
  end_if;

  //look for right Identifier
  if ( a_data[ 0 ] <> 16#12345678 ) then
    sd_retval := -102;
    return;
  end_if;

  //look for valid length	(we only read 128 Byte at the moment [16Byte are header])
  if( a_data[ 3 ] > (128 - 16 ) ) then
    sd_retval := -103;
    return;
  end_if;

  //search for SPI Flash Configuration
  for i := 0 to a_data[ 3 ] / sizeof( UDINT ) do

    //look for configuration id in 3rd byte
    if ( ( a_data[ i + 4 ] and 16#FF00_0000 ) = SearchID ) then
      p_BaseListAddress^ := a_data[ i + 4 ] and 16#00FF_FFFF;
      sd_retval := 0;
      return;
    end_if;

  end_for;

  //if no entry is found
  sd_retval := -100;

END_FUNCTION

FUNCTION VaranManager::GetDocuFileInfo
  VAR_INPUT
    p_us_position_info 	: ^USINT;
    ud_listOffset 	    : UDINT;
  END_VAR
  VAR_OUTPUT
    sd_retval 	        : DINT;
  END_VAR
  VAR
    a_data			        : ARRAY[0..2] OF UDINT;
  END_VAR

  //read header of documentation list
  sd_retval := ReadSPIDataComfort(p_us_position_info  := p_us_position_info,
                                  ud_offset           := ud_listOffset,
                                  ud_length	          := sizeof(a_data),
                                  p_data	            := ( #a_data )$^USINT
                                 );

  //look for an error
  if ( sd_retval <> VARANMANAGER_OK ) then
    return;
  end_if;

  // check if length is > 0
  if ( a_data[ 2 ] = 0 ) then
    sd_retval := -100;
    return;
  end_if;

  // save length of file
  ud_SPI_Docu_Length := a_data[ 2 ];

  //offset = listoffset + 4 byte for checksum + 4 byte for list version + 4 byte length
  ud_SPI_Offset := ud_listOffset + 12;

END_FUNCTION

FUNCTION VaranManager::ReadSPIDataComfort
  VAR_INPUT
    p_us_position_info 	: ^USINT;
    ud_offset 	        : UDINT;
    ud_length 	        : UDINT;
    p_data 	            : ^USINT;
  END_VAR
  VAR_OUTPUT
    sd_retval 	        : DINT;
  END_VAR
  VAR
    ud_read_length	    : UDINT;
  END_VAR

  //look if we have a length
  if ( ud_length = 0 ) then
    sd_retval := -100;
    return;
  end_if;

  //look if data is in one page
  while ( ud_length <> 0 ) do

    //if length is above page size
    if ( ( ud_offset and 16#FF ) + ud_length > 16#FF ) then
      //how many bytes are in this page available
      ud_read_length := 16#100 - ( ud_offset and 16#FF );
      //not more than 128 Bytes
      if ( ud_read_length > 128 ) then
        ud_read_length := 128;
      end_if;
    else
      //not more than 128 Bytes
      if ( ud_length > 128 ) then
        ud_read_length := 128;
      else
        ud_read_length := ud_length;
      end_if;
    end_if;

    //read data
    sd_retval :=      ReadSPIData( p_us_position_info	:= p_us_position_info,
                                   ud_offset				  := ud_offset,
                                   ud_length				  := ud_read_length,
                                   p_data				      := p_data
                                 );
    //look for an error
    if ( sd_retval <> VARANMANAGER_OK ) then
//			State := _SPIError;
      return;
    end_if;

    //correct length
    ud_length -= ud_read_length;
    ud_offset += ud_read_length;
    p_data    += ud_read_length;
  end_while;

END_FUNCTION

FUNCTION VIRTUAL GLOBAL VaranManager::GetSerialNo
  VAR_INPUT
    p_us_position_info 	: ^USINT;
    p_SerialNo 	        : ^CHAR;
  END_VAR
  VAR_OUTPUT
    sd_retval 	        : DINT;
  END_VAR
  VAR
    BaseListAddress     : UDINT;
    a_data              : ARRAY[0..31] OF UDINT;
  END_VAR

  if p_us_position_info & p_SerialNo then

    //check OS version
    if ( _RTOSVersion < VM_SPI_OS_VERSION ) then
      // access of SPI flash not possible
      sd_retval := -2;
      return;
    end_if;

    // check if documentation is available and get file size and offset in SPI flash
    if ( SearchSPIList(p_us_position_info, VM_SPI_SERIALNO_ID, #BaseListAddress) <> VARANMANAGER_OK ) then
      sd_retval := -3;
      return;
    end_if;

    //read header of serial number list
    sd_retval := ReadSPIDataComfort(p_us_position_info  := p_us_position_info,
                                    ud_offset           := BaseListAddress,
                                    ud_length	          := 12,
                                    p_data	            := ( #a_data )$^USINT
                                   );

    //look for an error and check if length is > 0
    if ( sd_retval <> VARANMANAGER_OK ) | ( a_data[ 2 ] = 0 ) then
      sd_retval := -4;
      return;
    end_if;

    //read the whole serial number string
    sd_retval := ReadSPIDataComfort( p_us_position_info := p_us_position_info,
                                     ud_offset	        := BaseListAddress + 12,
                                     ud_length	        := a_data[ 2 ],
                                     p_data		          := p_SerialNo
                                   );

    //add string termination
    (p_SerialNo + a_data[ 2 ])^ := 0;

    //look for an error
    if ( sd_retval <> VARANMANAGER_OK ) then
      sd_retval := -5;
      return;
    end_if;
  else
    // invalid parameters
    sd_retval := -1;
  end_if;

END_FUNCTION

FUNCTION VIRTUAL GLOBAL VaranManager::AllowRequiredError
  VAR_OUTPUT
    sd_retval 	: DINT;
  END_VAR

  SetRequiredError  := TRUE;
  sd_retval         := 0;

END_FUNCTION

FUNCTION VIRTUAL GLOBAL VaranManager::SetObjectThisp
  VAR_INPUT
    p_us_ObjectPath 	: ^USINT;
    ud_thisp 	        : UDINT;
  END_VAR
  VAR_OUTPUT
    sd_retval 	      : DINT;
  END_VAR

  if ( pHardwareTree <> NIL ) then
    sd_retval := HWT_iSetObjectThisp(VaranManagerNr,p_us_ObjectPath,ud_thisp);
  else
    sd_retval := 0;
  end_if;

END_FUNCTION

FUNCTION VIRTUAL GLOBAL VaranManager::GetObjectThisp
  VAR_INPUT
    p_us_ObjectPath : ^USINT;
  END_VAR
  VAR_OUTPUT
    ud_thisp 	      : UDINT;
  END_VAR

  if ( pHardwareTree <> NIL ) then
    ud_thisp := HWT_iGetObjectThisp(VaranManagerNr,p_us_ObjectPath);
  else
    ud_thisp := 0;
  end_if;

END_FUNCTION

//BLEERN001 start
FUNCTION VIRTUAL GLOBAL VaranManager::UpdateRtPostScan
VAR
  i                   : UDINT;
  pHelp               : ^t_s_OneHandle;
  AliveCheck          : DINT;
#ifndef VARAN_TIME_MEASUREMENT_DEACTIVATE
  ud_time	      	    : UDINT;
#endif
  ud_TempPllStatus    : UDINT;
#ifdef VARAN_TIME_MEASUREMENT_SINGLE_OBJECTS
  ud_SingleTimeMark1  : UDINT;
  ud_SingleTimeMark2  : UDINT;
#endif
END_VAR

  IF (us_RtStep <> _RtWork) THEN
    return;
  END_IF;

  if ManagerOn then

    //look if we have classes
    if ( s_RtPostScanHandles.ud_NrOfHandles > 0 ) then

      //call all connected classes
      pHelp := #s_RtPostScanHandles.p_HandleList^[0];
      for i := 0 to s_RtPostScanHandles.ud_NrOfHandles - 1 do

#ifdef VARAN_TIME_MEASUREMENT_SINGLE_OBJECTS
        ud_SingleTimeMark1 := OS_READMICROSEC();
#endif

        //call class
        pHelp^.p_This^.UpdateRtPostScan();

#ifdef VARAN_TIME_MEASUREMENT_SINGLE_OBJECTS
        ud_SingleTimeMark2 := OS_READMICROSEC();
        pHelp^.TimeMeasuring.ud_ActTime := ud_SingleTimeMark2 - ud_SingleTimeMark1;

        if pHelp^.TimeMeasuring.ud_ActTime > pHelp^.TimeMeasuring.ud_MaxTime then
          pHelp^.TimeMeasuring.ud_MaxTime := pHelp^.TimeMeasuring.ud_ActTime;
        end_if;

        if pHelp^.TimeMeasuring.ud_ActTime < pHelp^.TimeMeasuring.ud_MinTime then
          pHelp^.TimeMeasuring.ud_MinTime := pHelp^.TimeMeasuring.ud_ActTime;
        end_if;
#endif

        //get pointer on next handle
        pHelp += sizeof(t_s_OneHandle);
      end_for;
    end_if;

    if ( IsAlsoClient & p_ManagerClientSpace <> NIL ) then

      //increment alive counter
      pIsoWriteSafetyData^.VMC_Header.ui_AliveCounter += 1;

      if b_PayloadSupport &
         pMultiVaran^.udVersion >= VM_MULTIVARAN_VERSION_FULL_PAYLOAD_AVAILABLE  then
        MULTI_VARAN_iGetNodeProperty( hNodeHandle       := vmNodeHandle
                                    , udPropertyId      := VM_PROP_PLL_STATUS_REGISTER
                                    , pudPropertyValue  := #ud_TempPllStatus
                                    );
        pIsoWriteSafetyData^.VMC_Header.us_Status.PLL_Locked := (ud_TempPllStatus AND 2#0101) = 2#0101; // check pll locked and device delay time compensated bit
      else

        pIsoWriteSafetyData^.VMC_Header.us_Status.PLL_Locked := (p_ManagerPll^.ucControlStatus AND 2#0101) = 2#0101; // check pll locked and device delay time compensated bit
      end_if;

      if bPdoCopyDisable = false then

        // copy safety data from application memory to manager DPRAM
        if pIsoWriteSafetyData then
          To_Stdlib.MemCpy( dest    := p_ManagerClientSpace + VM_CLIENT_ISO_WR_OFFSET,
                            source  := pIsoWriteSafetyData,
                            size    := (SafetyIsoMemWrite + VM_CLIENT_HEADER_SIZE)$UDINT
                          );
        end_if;
      else
        // copy data from application memory
        if pIsoWriteSafetyData then
          // copy header and TDO data from application memory
          To_Stdlib.MemCpy( dest    := p_ManagerClientSpace + VM_CLIENT_ISO_WR_OFFSET
                          , source  := pIsoWriteSafetyData
                          , size    := sizeof(t_VMC_Header) + sizeof(t_VMC_Safety_Header_TDO)
                          );
        end_if;
      end_if;
      // copy user PDO data from application to manager DPRAM
      if UserObjectData.pIsoWriteData then
        To_Stdlib.MemCpy( dest    := p_ManagerClientSpace + VM_CLIENT_ISO_WR_OFFSET + SafetyIsoMemWrite + VM_CLIENT_HEADER_SIZE,
                          source  := UserObjectData.pIsoWriteData,
                          size    := UserObjectData.udIsoWriteLength
                        );
      end_if;

      //******************************************************************************************************

      // check AliveCounter every Xth cycle (because the other system may have a different speed)
      if pIsoWriteSafetyData^.VMC_Header.ui_AliveCounter MOD VMC_ModValue = 0 then
        //check alive counter
        AliveCheck := pIsoReadSafetyData^.VMC_Header.ui_AliveCounter - ui_AliveCounterOld;
        if ( AliveCheck$INT <= 0 ) then
          SyncCheck := 0;
        else
          SyncCheck := (SyncCheck SHL 1) OR pIsoWriteSafetyData^.VMC_Header.us_Status.PLL_Locked;
        end_if;
        ui_AliveCounterOld := pIsoReadSafetyData^.VMC_Header.ui_AliveCounter;

        if SyncCheck = 16#FF then
          SuperiorSystemOK  := 1;
          TriggerClientWD   := FALSE;
        else
          SuperiorSystemOK  := 0;
          UnSyncCounter     += 1;
        end_if;
      end_if;
    else
      SuperiorSystemOK := -1;
    end_if;

    ExecuteDOL( VARAN_DOL_ISO );

#ifndef VARAN_TIME_MEASUREMENT_DEACTIVATE
    //get rt time

    if b_PayloadSupport &
       pMultiVaran^.udVersion >= VM_MULTIVARAN_VERSION_FULL_PAYLOAD_AVAILABLE  then
      MULTI_VARAN_iGetTimeUpCounter( hManagerNodeHandle := vmNodeHandle
                                   , pudTimeUpCounterNs := #ud_time
                                   );
    else
      ud_time := p_ManagerStructure^.uiTUpCounter;
    end_if;

    //get call time
    s_VaranTimes.s_Realtime.ud_ActTime := Act_RtTime := ( ud_time - s_VaranTimes.s_Realtime.ud_Timemark ) / 1000;

    //look for maximum
    if ( Act_RtTime > Max_RtTime ) then
      Max_RtTime := Act_RtTime;
    end_if;

    //look for minimum
    if ( Act_RtTime < Min_RtTime ) then
      Min_RtTime := Act_RtTime;
    end_if;
#endif

  end_if;

END_FUNCTION

#pragma warning(disable:73)
FUNCTION GLOBAL VaranManager::TopologyChangeLogin
  VAR_INPUT
    pServer 	: ^DINT;
  END_VAR
#pragma warning(default:73)
// the whole method makes no sense, if we don't get a callback
#ifdef VARAN_iSetManagerCallbackOnConnect
  VAR
    pHelp     : ^t_s_FlexHub;
  END_VAR

  // general callback works only on os versions >= 01.02.085
  if _RTOSVersion >= 16#1255 then
    if pFlexHubs = NIL then
      pFlexHubs$pVoid := To_StdLib.Malloc(size:=sizeof(t_s_FlexHub));
      pHelp := pFlexHubs;

      // if there is no VARAN Interface available, we would crash at the call
      if pVaran = NIL then
        return;
      end_if;

      // only on the first login we call the OS interface
      VARAN_iSetManagerCallbackOnConnect(1);
    else
      pHelp := pFlexHubs;
      while pHelp^.pNext <> NIL do
        pHelp := pHelp^.pNext;
      end_while;
      pHelp^.pNext$pVoid := To_StdLib.Malloc(size:=sizeof(t_s_FlexHub));
      pHelp := pHelp^.pNext;
    end_if;

    if pHelp <> NIL then
      pHelp^.pServer := pServer - sizeof(SvrCh.pMeth);
      pHelp^.pNext   := NIL;
    end_if;
  else

#ifdef HWC_LogError
    HWC_LogError(this,"@019B (VaranManager::TopologyChangeLogin) General callback for FlexHub works only on os versions >= 01.02.085");
#endif

  end_if;
#else
#ifdef HWC_LogError
 HWC_LogError(this,"@019C (VaranManager::TopologyChangeLogin) Need newer lsl_st_varan.h file for general callback functionality");
#endif
  #pragma message("Need newer lsl_st_varan.h file for general callback functionality (used for FlexHub class)")
#endif

END_FUNCTION

FUNCTION GLOBAL VaranManager::AddDAClientRdData
  VAR_INPUT
    ud_length 	: UDINT;
    p_pdata 	  : ^void;
    pThis 	    : ^void;
    pFunction 	: ^void;
  END_VAR
  VAR_OUTPUT
    sd_retval 	: DINT;
  END_VAR

  //check if manager is also client
  if (IsAlsoClient = 0) | (SuperiorSystemTime = 0) then
    sd_retval := -6;
    return;
  end_if;

  //check length (we reserve 4 bytes for header)
  if ( ud_length > (VM_CLIENT_MAX_BUFFER_USE - VM_CLIENT_HEADER_SIZE) ) then
    sd_retval := -2;
    return;
  end_if;

  //check pointer
  if ( p_pdata = NIL ) | (pThis = NIL) | (pFunction = NIL) then
    sd_retval := -3;
    return;
  end_if;

  // check fpga version (must be >= 1.4) and os version (must be >= 01.02.103)
  if Release < 16#14 then

    // fpga doesn't support the new buffer
    sd_retval := -7;
#ifdef HWC_LogError
    HWC_LogError(this, "@019D (VaranManager::AddDAClientRdData) FPGA version of VMC needs to be at least 1.4 to support the direct access buffer");
#endif
    return;

  elsif _RTOSVersion < VM_DA_BUFFER_AVAILABLE then

    // os doesn't support the irq callback
    sd_retval := -8;
#ifdef HWC_LogError
    HWC_LogError(this, "@019E (VaranManager::AddDAClientRdData) For IRQ Callback on VMC buffer os version >= 01.02.103 is required");
#endif
    return;
  else

#ifdef VARAN_iSetManagerCallbackOnVmcBufDaInt
    // if there is no VARAN Interface available, we would crash at the call
    if pVaran = NIL then
      sd_retval := VARANMANAGER_DRIVER_NOT_EXISTS;
      return;
    end_if;

    // install irq callback
    VARAN_iSetManagerCallbackOnVmcBufDaInt(1);
    DA_IRQ_pFunc  := pFunction;
    DA_IRQ_pthis  := pThis;

    //save length and data pointer
    DA_IRQ_Length := ud_length ;
    DA_IRQ_pData  := p_pdata;

#else
    // newer lsl_st_varan.h neccessary to use this functionality
    sd_retval := -9;
#ifdef HWC_LogError
    HWC_LogError(this, "@019F (VaranManager::AddDAClientRdData) Need newer lsl_st_varan.h file to install IRQ Callback on VMC direct access buffer");
#endif
    #pragma message("Need newer lsl_st_varan.h file to install IRQ Callback on VMC direct access buffer");
    return;
#endif
  end_if;

  sd_retval := 0;

END_FUNCTION

FUNCTION GLOBAL VaranManager::SendDAClientWrData
  VAR_INPUT
    ud_length 	: UDINT;
    p_pdata 	  : ^void;
  END_VAR
  VAR_OUTPUT
    sd_retval 	: DINT;
  END_VAR

  //check if manager is also client
  if (IsAlsoClient = 0) | (SuperiorSystemTime = 0) then
    sd_retval := -6;
    return;
  end_if;

  //check support of da buffer
  if Release < 16#14 then
    sd_retval := -1;
    return;
  end_if;

  //check length (we reserve 4 bytes for header)
  if ( ud_length > (VM_CLIENT_MAX_BUFFER_USE - VM_CLIENT_HEADER_SIZE) ) then
    sd_retval := -2;
    return;
  end_if;

  //check pointer
  if ( p_pdata = NIL ) then
    sd_retval := -3;
    return;
  end_if;

  // save data to output data memory
  if ud_length > VM_CLIENT_HEADER_SIZE then
    To_Stdlib.MemCpy(dest   := p_ManagerClientSpace + VM_CLIENT_DA_WR_OFFSET + VM_CLIENT_HEADER_SIZE
                   , source := p_pdata + VM_CLIENT_HEADER_SIZE
                   , size   := ud_length - VM_CLIENT_HEADER_SIZE
                   );
  end_if;

  // the first 4 byte are written in the end (switch buffer)
  (p_ManagerClientSpace + VM_CLIENT_DA_WR_OFFSET)^ := p_pdata^$DINT;

  sd_retval := 0;

END_FUNCTION

FUNCTION VIRTUAL GLOBAL VaranManager::GetNsTimeBPLLTicks
  VAR_OUTPUT
    ud_ns_counter 	: UDINT;
  END_VAR

  //look if init has been executed
  if ( s_VaranManagerSettings.us_InitCounter = 0 ) then
    bExternalInit := true;
    Init();
  end_if;

  if b_PayloadSupport &
    pMultiVaran^.udVersion >= VM_MULTIVARAN_VERSION_FULL_PAYLOAD_AVAILABLE  then
    MULTI_VARAN_iGetNodeProperty( hNodeHandle       := vmNodeHandle
                                , udPropertyId      := VM_PROP_TIME_UP_COUNTER_BETWEEN_PLL_TICKS
                                , pudPropertyValue  := #ud_ns_counter
                                );
  else

    //if we have the Manager structure
    if ( p_ManagerStructure <> NIL ) then
      ud_ns_counter := p_ManagerStructure^.uiTUpCounterBPLLTicks;
    end_if;
  end_if;

END_FUNCTION

FUNCTION VIRTUAL GLOBAL VaranManager::AddMovDO
  VAR_INPUT
    ud_dol_type 	      : UDINT;
    p_ud_handle 	      : ^UDINT;
    p_ud_MovSettings 	  : ^UDINT;
    ud_type 	          : UDINT;
  END_VAR
  VAR_OUTPUT
    sd_retval 	        : DINT;
  END_VAR
  VAR
    p_dummy             : UDINT;
    pVaranHandle        : ^LSL_VARANFRAME;
//    TempMem             :  UDINT;
  END_VAR

#ifdef VM_DEBUG_PAYLOAD
  // Payload not supported
  if b_PayloadSupport then
    // This method is not supporded with Payload support
    ((0)$^USINT)^ := 0;
  end_if;
#endif

  if p_ud_MovSettings then

    // add data object Move Command (add write and change the command type)
    sd_retval := AddWrDO( p_us_position_info:=NIL
                        , ud_dol_type:=ud_dol_type
                        , p_ud_handle:=p_ud_handle
                        , ud_address:=0
                        , ud_length:=0
                        , p_ud_data:= #p_dummy
                        , ud_type:= VM_MEMORY_ACCESS
                        );

    // if no error, we initialize the return structure
    if ( sd_retval = VARANMANAGER_OK ) then
      // check if the DO has a special priority
      if ud_type AND VM_PRIORITY_FILTER then
        AddToDOPriorityList(p_ud_handle^$^LSL_VARANFRAME, ud_type AND VM_PRIORITY_FILTER);
      end_if;

      pVaranHandle              := (p_ud_handle^)$^LSL_VARANFRAME;

      // replace the write command with the move command
      pVaranHandle^.ucDOType    := 16#10;

      // start with not moving anything
      pVaranHandle^.ucCtrlStat  := VARAN_DO_NO_RUN;

      // start of the mover settings is, where normally the ucRetrys is (no retries necessary in local memory)
      p_ud_MovSettings^         := (#pVaranHandle^.ucRetrys)$UDINT;

(*    // is already counted with the AddWrDO-Call
      //26 Byte (Header) + 2 Byte (compensate missalignment)
      TempMem := 28;

      case ud_dol_type of
      // **************************************************
        VARAN_DOL_DA:
          DPRAM_Used.DA_RdWr += TempMem;
          DOCounter.DA_RdWr  += 1;
      // **************************************************
        VARAN_DOL_ISO:
          DPRAM_Used.ISO_RdWr += TempMem;
          DOCounter.ISO_RdWr  += 1;
      // **************************************************
        VARAN_DOL_ASY:
          DPRAM_Used.ASY_RdWr += TempMem;
          DOCounter.ASY_RdWr  += 1;
      // **************************************************
        VARAN_DOL_ADMIN:
          DPRAM_Used.Admin_RdWr += TempMem;
          DOCounter.Admin_RdWr  += 1;
      // **************************************************
        VARAN_DOL_IRQ:
          DPRAM_Used.IRQ_RdWr += TempMem;
          DOCounter.IRQ_RdWr  += 1;
      end_case;
*)
    else
      p_ud_MovSettings^ := NIL;
    end_if;

  end_if;

END_FUNCTION

// Method not used with Payload DO's, OS Handles priority's in this case.
FUNCTION VaranManager::AddToDOPriorityList
  VAR_INPUT
    pHandle 	    : ^LSL_VARANFRAME;
    ud_Priority 	: HDINT;
  END_VAR
  VAR
    pListHelp     : ^t_PrioListList;
    pHelp         : ^t_PrioHandleList;
  END_VAR

  // if there is no VARAN Interface available, we would crash at adding dummy DOs
  if pVaran = NIL then
    return;
  end_if;

  // check if there is already a list with a priority
  if pPriorityList = NIL then
    // if not, create it
    pPriorityList$pVoid := To_StdLib.Malloc(size:=sizeof(t_PrioListList));
    pListHelp := pPriorityList;
    if pListHelp <> NIL then
      pListHelp^.Prio  := ud_Priority;
      pListHelp^.pList := NIL;
      pListHelp^.pNext := NIL;
    else
      // failed to allocate memory
      State := _NoMem;
      return;
    end_if;
  else
    pListHelp := pPriorityList;
    while (pListHelp^.Prio <> ud_Priority) & (pListHelp^.pNext <> NIL) do
      pListHelp := pListHelp^.pNext;
    end_while;
    if (pListHelp^.Prio <> ud_Priority) then
      pListHelp^.pNext$pVoid := To_StdLib.Malloc(size:=sizeof(t_PrioListList));
      pListHelp := pListHelp^.pNext;
      if pListHelp <> NIL then
        pListHelp^.Prio  := ud_Priority;
        pListHelp^.pList := NIL;
        pListHelp^.pNext := NIL;
      else
        // failed to allocate memory
        State := _NoMem;
        return;
      end_if;
    end_if;
  end_if;

  // now we have the pointer to the list of the right priority (pListHelp^.pList)

  // check if there is already an entry with this handle
  if pListHelp^.pList = NIL then
    // if not, create it
    pListHelp^.pList$pVoid := To_StdLib.Malloc(size:=sizeof(t_PrioHandleList));
    pHelp := pListHelp^.pList;
  else
    pHelp := pListHelp^.pList;
    while (pHelp^.pHandle <> pHandle) & (pHelp^.pNext <> NIL) do
      pHelp := pHelp^.pNext;
    end_while;
    if (pHelp^.pHandle <> pHandle) then
      pHelp^.pNext$pVoid := To_StdLib.Malloc(size:=sizeof(t_PrioHandleList));
      pHelp := pHelp^.pNext;
    else
      // already in list
      return;
    end_if;
  end_if;

  if pHelp <> NIL then
    pHelp^.pHandle := pHandle;
    pHelp^.pNext := NIL;
  else
    // failed to allocate memory
    State := _NoMem;
    return;
  end_if;

END_FUNCTION

// Method not used with Payload DO's, OS Handles priority's in this case.
FUNCTION VaranManager::SortCmdsByPriority
  VAR
    pHelpFrame        : ^LSL_VARANFRAME;
    pHelp             : ^t_PrioHandleList;
    pNonPrioList      : ^t_PrioHandleList;
    pActList          : ^t_PrioListList;
    pNextList         : ^t_PrioListList;
    pPreviousList     : ^t_PrioListList;
    bMadeSort         : BOOL;
    sd_retval         : DINT;
    pDummyReadData    : UDINT;
    pDummyHandle      : UDINT;
    pTerminationFrame : ^LSL_VARANFRAME;
  END_VAR

  // search for first command which is not in priority list
  pHelpFrame := p_SyncAndWdDO;

  // if first command is not sync, we don't sort anything (check command = 0 and subcommand = 1) => some error may have occured
  if ((((#pHelpFrame^.uiResponseTime)$^USINT + 4)^ AND 16#F0) = 0) & (((#pHelpFrame^.uiResponseTime)$^USINT + 5)^ = 1) then

    // add a dummy DO just to be the last one after sorting (otherwise the OS can't add DOs during runtime like for DIAS DRIVE)
#pragma warning(disable: 75)
    sd_retval := VARAN_iAddDOToDOL	( uiManager			  := VaranManagerNr
                                    , pucNode			    := NIL
                                    , uiDOLType 		  := VARAN_DOL_ISO
                                    , puiDOHandle		  := #pDummyHandle
                                    , uiCmd				    := VARAN_CMD_MEMORY_READ
                                    , uiAddressRead		:= 0
                                    , uiLengthRead		:= 1
                                    , pucRead			    := #pDummyReadData
                                    , uiAddressWrite	:= 0
                                    , uiLengthWrite		:= 0
                                    , pucWrite			  := NIL
                                    );
#pragma warning(default: 75)

    //if an error occured => we don't sort anything
    if ( sd_retval <> VARANMANAGER_OK ) then
      // tell the RT that we're finished with sorting
      us_RtStep := _Wait4Sync;
      return;
    end_if;

    pNonPrioList  := NIL;
    pHelpFrame    := pHelpFrame^.pNext$^LSL_VARANFRAME;
    while pHelpFrame <> 16#FFFFFFFF do

      if IsInPriorityList(pHelpFrame) = FALSE then
        // put the non-priored commands in an own list (without sync)

        if pNonPrioList = NIL then
          // if not, create it
          pNonPrioList$pVoid := To_StdLib.Malloc(size:=sizeof(t_PrioHandleList));
          pHelp := pNonPrioList;
        else
          pHelp := pNonPrioList;
          while (pHelp^.pNext <> NIL) do
            pHelp := pHelp^.pNext;
          end_while;
          pHelp^.pNext$pVoid := To_StdLib.Malloc(size:=sizeof(t_PrioHandleList));
          pHelp := pHelp^.pNext;
        end_if;

        if pHelp <> NIL then
          pHelp^.pHandle := pHelpFrame;
          pHelp^.pNext := NIL;
        else
          // failed to allocate memory
          State := _NoMem;
          return;
        end_if;
      end_if;

      if pHelpFrame^.pNext = 16#FFFFFFFF then
        pTerminationFrame := pHelpFrame;
      end_if;

      pHelpFrame := pHelpFrame^.pNext$^LSL_VARANFRAME;
    end_while;

    // now we got the priorized and the non-priorized commands

    // sort the lists by priority number
    bMadeSort := TRUE;
    while bMadeSort do
      bMadeSort := FALSE;

      // go through all priority lists
      pPreviousList := pActList := pPriorityList;
      while pActList^.pNext do
        // if the next list has a higher priority number => resort it
        if pActList^.Prio > pActList^.pNext^.Prio then
          pNextList         := pActList^.pNext;

          pActList^.pNext   := pNextList^.pNext;
          pNextList^.pNext  := pActList;

          // if it's the first module, we have to change also the pointer to the list
          if pPriorityList = pActList then
            pPreviousList         := pPriorityList := pNextList;
          else
            // if the beginning of the list has changed it doesn't count, because then we start again automatically
            bMadeSort             := TRUE;
            pPreviousList^.pNext  := pNextList;
          end_if;
          pActList := pNextList;
        else
          pActList := pActList^.pNext;
        end_if;

        if (pActList <> pPriorityList) & (pActList <> pPriorityList^.pNext) then
          pPreviousList := pPreviousList^.pNext;
        end_if;
      end_while;
    end_while;

    // the lists in pPriorityList are now sorted by priority => hang the non-priorized list as last priority after this
    pActList := pPriorityList;
    while (pActList^.pNext <> NIL) do
      pActList := pActList^.pNext;
    end_while;
    pActList^.pNext$pVoid := To_StdLib.Malloc(size:=sizeof(t_PrioListList));
    pActList := pActList^.pNext;
    if pActList <> NIL then
      pActList^.Prio  := 16#FFFFFFFF;
      pActList^.pList := pNonPrioList;
      pActList^.pNext := NIL;
      pNonPrioList    := NIL;  // no more need to remember this
    else
      // failed to allocate memory
      State := _NoMem;
      return;
    end_if;

    // change pNext of Sync-Command to the first command of our list
    p_SyncAndWdDO^.pNext$^LSL_VARANFRAME := pPriorityList^.pList^.pHandle;

    // and now we go through the list and change all next pointers (priority is automatically given)
    pActList := pPriorityList;
    while pActList do
      // go through all elements of this list
      pHelp := pActList^.pList;
      while pHelp^.pNext do
        pHelp^.pHandle^.pNext$^LSL_VARANFRAME := pHelp^.pNext^.pHandle;

        pHelp := pHelp^.pNext;
      end_while;

      if pActList^.pNext then
        pHelp^.pHandle^.pNext$^LSL_VARANFRAME := pActList^.pNext^.pList^.pHandle;
      end_if;

      pActList := pActList^.pNext;
    end_while;
  end_if;

END_FUNCTION

// Method not used with Payload DO's, OS Handles priority's in this case.
FUNCTION VaranManager::IsInPriorityList
  VAR_INPUT
    pHandle 	: ^LSL_VARANFRAME;
  END_VAR
  VAR_OUTPUT
    retcode 	: BOOL;
  END_VAR
  VAR
    pListHelp : ^t_PrioListList;
    pHelp     : ^t_PrioHandleList;
  END_VAR

  retcode := FALSE;

  // go through all priority lists
  pListHelp := pPriorityList;
  while pListHelp do
    // go through all elements of this list
    pHelp := pListHelp^.pList;
    while pHelp do
      // check if it's the handle we search for
      if pHelp^.pHandle = pHandle then
        retcode := TRUE;
        return;
      end_if;

      pHelp := pHelp^.pNext;
    end_while;

    pListHelp := pListHelp^.pNext;
  end_while;

END_FUNCTION

FUNCTION VaranManager::FirstInit
VAR
  sd_retval     	    : DINT;
  ud_counter	        : UDINT;
  i		          	    : UDINT;
  ManagerNodeString   : USINT;
  nodeProperty        : ARRAY [0..2] of LSL_PROPERTY_VALUE_PAIR;
  aStrSemaphore       : ARRAY [0..99] of CHAR;
  aStrVaranManagerNr  : ARRAY [0..5] of CHAR;
  udTempCyTime        : UDINT;
END_VAR

  bFirstInitDone      := true;

  //read Clients
  VaranManagerNr	    := VaranManagerNr.read();
  VaranManagerTime    := VaranManagerTime.read();
//  IRQTaskTime         := IRQTaskTime.read();
  IsAlsoClient        := IsAlsoClient.read();
  SuperiorSystemTime  := SuperiorSystemTime.Read();

  //Check if varanmanager number is available on HW
  if VaranManagerNr > udSystemVaranManagerCnt then
#ifdef HWC_LogError
    HWC_LogValue2(this, "@01A0 (VaranManager::FirstInit) Invalid varanmanagernumber 0x{0}! Max. number on this CPU is 0x{1}", VaranManagerNr ,udSystemVaranManagerCnt);
#endif
    state := _ManagerError;
    ManagerOn := 0;
    return;
  end_if;

  //set limit for VaranManagerTime
  if VaranManagerTime > 32000000 then
#ifdef HWC_LogError
    HWC_LogError(this, "@0026 (VaranManager::FirstInit) Maximum limit for VaranManagerTime (32 000 000 ns = 32 ms) exceeded");
#endif
    state := _VaranTimeError;
    ManagerOn := 0;
    return;
  end_if;

  //get rt-debug state
  b_RtDebug := To_HwControl.GetRtDebugState() <> 0;

  //****************************************************************************
  if b_PayloadSupport
     & pMultiVaran^.udVersion >= VM_MULTIVARAN_DOL_SET_REQUIRED_ERROR_ISO_START_TIME then

    //-----------------------------------------------------------------------------------------------
    //get manager node info from os
    p_NodeInfo := #s_NodeInfo;

    sd_retval := MULTI_VARAN_iGetNodeInformation( hNodeHandle := vmNodeHandle
                                                , psNodeInfo  := p_NodeInfo
                                                );

    if	( sd_retval <> VARANMANAGER_OK
      | p_NodeInfo = NIL
      )
    then
      State := _NoHardware;
      return;
    end_if;

    // get release of FPGA
    Release := p_NodeInfo^.ucFPGAVersion;

  //-----------------------------------------------------------------------------------------------

    p_SyncOut := #s_SyncOut;

    // disable varan manager sync out
    // Searching for the correct sync is no longer nessersary because we pass the sync ID when it is configured
    // The value will be writted o the VM later in this method with MULTI_VARAN_ICONFIGUREPLLSYNCOUT
    p_SyncOut^.ucControlStatus      := 0;

    // set required bit on (for varan error in init (os set bit in function InitApp) later)
    nodeProperty[0].udPropertyId    := VM_PROP_REQUIRED_ERROR_ENABLED;
    nodeProperty[0].udPropertyValue := 1;
    MULTI_VARAN_iSetNodeProperties( hNodeHandle           := vmNodeHandle
                                  , udPropertyCount       := 1
                                  , psPropertyValuePairs  := #nodeProperty[0]
                                  );

    //Get ISO start Time
    GetISOStartTime();

    s_ManagerControlData.ud_IsoStartPoint := VaranManagerTime * IsoStartPoint / 100;

    nodeProperty[0].udPropertyId          := VM_PROP_ISO_START_TIME;
    nodeProperty[0].udPropertyValue       := s_ManagerControlData.ud_IsoStartPoint;
    MULTI_VARAN_iSetNodeProperties( hNodeHandle           := vmNodeHandle
                                  , udPropertyCount       := 1
                                  , psPropertyValuePairs  := #nodeProperty[0]
                                  );

    //Check if OS supports full payload
    if b_PayloadSupport &
       pMultiVaran^.udVersion < VM_MULTIVARAN_VERSION_FULL_PAYLOAD_AVAILABLE then

      //OS do not support full payload with the multivaran interface
      //so we need to use some functions from the old interface.

      //-----------------------------------------------------------------------------------------------
      //get Manager structure
      sd_retval := VARAN_iGetManagerControl	( uiManager := VaranManagerNr
                                            , pvCB 		  := ( #p_ManagerStructure )$^PLSL_CONTROLBLOCK
                                            , pvPLL		  := ( #p_ManagerPll )$^PLSL_VARANPLL
                                            );

      //look for an error
      if	( sd_retval 			<> 	VARANMANAGER_OK
        | p_ManagerStructure	=	NIL
        | p_ManagerPll			  =	NIL
        )
      then
        State 		:= _NotInitialized;
        ManagerOn	:= 0;
        return;
      end_if;

      //look for right sync out pointer
      p_SyncOut := #p_ManagerPll^.sSynOutPeripheral1;
      ud_Counter := VaranManagerNr;

      //look in all peripheral sync outs
      for i := 1 to VM_MAX_SYNC_OUTS - 1 do

        //look if sync out id is correct
        if ( p_SyncOut^.ucSyncOutID = VM_SYNC_OUT_ID ) then

          //if it is right pll for right manager number (first is vor VaranManager number 0, second for VaranManager number 1, ....)
          if ( ud_counter = 0 ) then
            exit;					//we found right sync out --> exit
          end_if;
          ud_counter -= 1;			//we find one for lower VaranManager number
        end_if;

        //get pointer to next sync out
        p_SyncOut += sizeof ( LSL_VARANPLLSYNCOUT );

        //if we searched all sync outs set VaranManager off
        if ( i = VM_MAX_SYNC_OUTS - 1 ) then
          p_SyncOut := NIL;
          State 		:= _NotInitialized;
          ManagerOn	:= 0;
          return;
        end_if;
      end_for;

      //disable varan manager sync out
      p_SyncOut^.ucControlStatus := 0;
    end_if;

  else // if b_PayloadSupport ****************************************************************************

    // if there is no VARAN Interface available, we would crash at the call
    if pVaran = NIL then
      sd_retval := VARANMANAGER_DRIVER_NOT_EXISTS;
      return;
    end_if;

      //-----------------------------------------------------------------------------------------------
    //get manager node info from os
    ManagerNodeString := 0;

    //call OS - function (must be OS-funciton because of error handling)
    sd_retval := VARAN_iGetNodeInfo	( uiManager	:= VaranManagerNr
                                    , pucNode	  := #ManagerNodeString
                                    , pNodeInfo	:= #p_NodeInfo
                                    );

    if	( sd_retval <> VARANMANAGER_OK
      | p_NodeInfo = NIL
      )
    then
      State := _NoHardware;
      return;
    end_if;

      // get release of FPGA
    Release := p_NodeInfo^.ucFPGAVersion;

    //-----------------------------------------------------------------------------------------------
    //get Manager structure
    sd_retval := VARAN_iGetManagerControl	( uiManager := VaranManagerNr
                                          , pvCB 		  := ( #p_ManagerStructure )$^PLSL_CONTROLBLOCK
                                          , pvPLL		  := ( #p_ManagerPll )$^PLSL_VARANPLL
                                          );

    //look for an error
    if	( sd_retval 			<> 	VARANMANAGER_OK
      | p_ManagerStructure	=	NIL
      | p_ManagerPll			= 	NIL
      )
    then
      State 		:= _NotInitialized;
      ManagerOn	:= 0;
      return;
    end_if;

    //look for right sync out pointer
    p_SyncOut := #p_ManagerPll^.sSynOutPeripheral1;
    ud_Counter := VaranManagerNr;

    //look in all peripheral sync outs
    for i := 1 to VM_MAX_SYNC_OUTS - 1 do

      //look if sync out id is correct
      if ( p_SyncOut^.ucSyncOutID = VM_SYNC_OUT_ID ) then

        //if it is right pll for right manager number (first is for VaranManager number 0, second for VaranManager number 1, ....)
        if ( ud_counter = 0 ) then
          exit;					//we found right sync out --> exit
        end_if;
        ud_counter -= 1;			//we find one for lower VaranManager number
      end_if;

      //get pointer to next sync out
      p_SyncOut += sizeof ( LSL_VARANPLLSYNCOUT );

      //if we searched all sync outs set VaranManager off
      if ( i = VM_MAX_SYNC_OUTS - 1 ) then
        p_SyncOut := NIL;
        State 		:= _NotInitialized;
        ManagerOn	:= 0;
        return;
      end_if;
    end_for;

    //disable varan manager sync out
    p_SyncOut^.ucControlStatus := 0;

    //set required bit on (for varan error in init (os set bit in function InitApp) later)
    p_ManagerStructure^.ucTCEnable := p_ManagerStructure^.ucTCEnable or 16#80;

    //Get ISO start Time
    GetISOStartTime();

    p_ManagerStructure^.uiIsoStartPoint := VaranManagerTime * IsoStartPoint / 100;

  end_if; // if b_PayloadSupport ****************************************************************************

  // get maintimer in ns to compare with varan times
  MainTimer := _ClockTicks * 1000;

  //look if VaranManagerTime is a multiple of maintimer (maintimer has to be always less or equal the varan time)
  if ( VaranManagerTime mod MainTimer <> 0 ) then
    //Log entry
#ifdef HWC_LogValue2
    HWC_LogValue2(this, "@064A (VaranManager::FirstInit) VaranManagerTime ({0}) is not a multiple of MainTimer ({1})!", VaranManagerTime, MainTimer);
#endif

    State 		:= _NotInitialized;
    ManagerOn	:= 0;
    return;
  end_if;

//------------------------------------------------------------ Client Instructions --------------------------------------------------------|
//                                                                                                                                         V
  if ( IsAlsoClient ) then

    if b_PayloadSupport &
       pMultiVaran^.udVersion >= VM_MULTIVARAN_VERSION_FULL_PAYLOAD_AVAILABLE  then
      sd_retval := MULTI_VARAN_iGetNodeProperty(  hNodeHandle       := vmNodeHandle
                                                , udPropertyId      := VC_OPT_PROP_BUFFER_ADDRESS_ISO // = Offset 0 in p_ManagerClientSpace
                                                , pudPropertyValue  := (#p_ManagerClientSpace)$^UDINT );

    elsif ( _RTOSVersion >= 16#11DA ) & pVaran then

      //Schnittstelle vom OS holen!!!!!!
      sd_retval := VARAN_iGetManagerClientAddress	( uiManager		:= VaranManagerNr
                                                  , uiType		  := 0
                                                  , puiAddress	:= ( #p_ManagerClientSpace )$^UDINT
                                                  );
    end_if;

    //check if function is available
    if ( sd_retval <> VARANMANAGER_OK | p_ManagerClientSpace = NIL ) then

      IsAlsoClient := 0;

#ifdef HWC_LogError
      HWC_LogError(this, "@0654 (VaranManager::FirstInit) Client - Function not available but activated! (at least OS - Version 1.1.217 required)");
#endif
    else
      TriggerClientWD             := TRUE;
      bEnableManagerWithNoModules := TRUE; // activate, to ensure varan-client functionality if no varan clients are connected to the manager.
      sd_retval                   := InitMulDivVMC();

      //look for an error
      if ( sd_retval <> 0 ) then
        ManagerOn	:= 0;
        return;
      end_if;
    end_if;

  end_if;

//------------------------------------------------------------ Client Instructions --------------------------------------------------------^
//                                                                                                                                         |

  //get system periode time
  if b_PayloadSupport &
     pMultiVaran^.udVersion >= VM_MULTIVARAN_VERSION_FULL_PAYLOAD_AVAILABLE  then

    if MULTI_VARAN_iGetNodeProperty( hNodeHandle       := vmNodeHandle
                                , udPropertyId      := VM_PROP_PLL_SYSTEM_PERIOD_TIME
                                , pudPropertyValue  := #ud_SystemPeriod
                                ) <> VARANMANAGER_OK then

#ifdef HWC_LogError
      HWC_LogError(this,"@01A1 (VaranManager::FirstInit) Failed to get PLL System period time");
#endif
